Fanuc KAREL source: KA00153.KL

PROGRAM KA00153
%NOLOCKGROUP
VAR
  SRC: ARRAY[4] OF INTEGER
  DST: ARRAY[4] OF JOINTPOS
BEGIN
  DST = SRC
END KA00153
